{attribute 'linkalways'} 
{attribute 'no_explicit_call' := 'This FB is a CLASS and must be accessed using methods or properties'}
{attribute 'enable_dynamic_creation'}
FUNCTION_BLOCK _ETcVnWorldCoordinateSystem EXTENDS EnumDatatypeBase
VAR
	localData : ETcVnWorldCoordinateSystem;
	activeData : REFERENCE TO ETcVnWorldCoordinateSystem;
	enumBaseDatatype : _DINT(localData);
END_VAR

METHOD PRIVATE AddLocalEnumeration
VAR_INPUT
	Enumeration : T_MAXSTRING;
	Value : ETcVnWorldCoordinateSystem;
END_VAR
AddEnumeration(Enumeration, Value);
END_METHOD

PROPERTY PUBLIC Address : PVOID
GET
Address := ADR(activeData);
END_GET
END_PROPERTY

METHOD PUBLIC ClearReference
VAR_INPUT
END_VAR
activeData REF= localData;
SetBaseDatatypeReference();
END_METHOD

METHOD PUBLIC Clone : I_Datatype
VAR
    pClone : POINTER TO _ETcVnWorldCoordinateSystem;
END_VAR
pClone := __NEW(_ETcVnWorldCoordinateSystem(InitialValue := Value));
Clone := pClone^;
END_METHOD

METHOD FB_init : BOOL
VAR_INPUT
	bInitRetains : BOOL; // if TRUE, the retain variables are initialized (warm start / cold start)
	bInCopyCode : BOOL;  // if TRUE, the instance afterwards gets moved into the copy code (online change)
	InitialValue : ETcVnWorldCoordinateSystem;
END_VAR
localData := InitialValue;
AddBaseDatatype(enumBaseDatatype);
ClearReference();

AddLocalEnumeration('TCVN_WCS_X_RIGHT_Y_DOWN' , ETcVnWorldCoordinateSystem.TCVN_WCS_X_RIGHT_Y_DOWN);
AddLocalEnumeration('TCVN_WCS_X_DOWN_Y_RIGHT', ETcVnWorldCoordinateSystem.TCVN_WCS_X_DOWN_Y_RIGHT);
AddLocalEnumeration('TCVN_WCS_X_LEFT_Y_DOWN', ETcVnWorldCoordinateSystem.TCVN_WCS_X_LEFT_Y_DOWN);
AddLocalEnumeration('TCVN_WCS_X_UP_Y_RIGHT', ETcVnWorldCoordinateSystem.TCVN_WCS_X_UP_Y_RIGHT);
AddLocalEnumeration('TCVN_WCS_X_RIGHT_Y_UP', ETcVnWorldCoordinateSystem.TCVN_WCS_X_RIGHT_Y_UP);
AddLocalEnumeration('TCVN_WCS_X_DOWN_Y_LEFT', ETcVnWorldCoordinateSystem.TCVN_WCS_X_DOWN_Y_LEFT);
AddLocalEnumeration('TCVN_WCS_X_LEFT_Y_UP', ETcVnWorldCoordinateSystem.TCVN_WCS_X_LEFT_Y_UP);
AddLocalEnumeration('TCVN_WCS_X_UP_Y_LEFT', ETcVnWorldCoordinateSystem.TCVN_WCS_X_UP_Y_LEFT);
END_METHOD

PROPERTY PUBLIC Identifier : T_MAXSTRING
GET
Identifier := 'ETcVnWorldCoordinateSystem';
END_GET
END_PROPERTY

METHOD IsEnumeratorValueEqual : BOOL
VAR_INPUT
	Enumerator : I_KeyValueForwardEnumerator;
END_VAR
VAR
	storedValue : ETcVnWorldCoordinateSystem;
END_VAR
IF NOT Enumerator.TryGet(storedValue) THEN
	RETURN;
END_IF

IsEnumeratorValueEqual := storedValue = activeData;
END_METHOD

METHOD PUBLIC MakeReferenceTo
VAR_INPUT
	ReferenceTarget : REFERENCE TO ETcVnWorldCoordinateSystem;
END_VAR
activeData REF= ReferenceTarget;
SetBaseDatatypeReference();
END_METHOD

METHOD PROTECTED SetBaseDatatypeReference
VAR_INPUT
END_VAR
enumBaseDatatype.MakeReferenceTo(activeData);
END_METHOD

PROPERTY PUBLIC Size : UDINT
GET
Size := SIZEOF(activeData);
END_GET
END_PROPERTY

METHOD TryMakeReferenceTo : BOOL
VAR_INPUT
	Target : I_Datatype;
END_VAR
VAR
	pTargetData : POINTER TO ETcVnWorldCoordinateSystem;
END_VAR
IF NOT IsEquivalentTo(Target) THEN
	RETURN;
END_IF

pTargetData := Target.Address;
activeData REF= pTargetData^;
SetBaseDatatypeReference();
TryMakeReferenceTo := TRUE;
END_METHOD

PROPERTY PUBLIC Value : ETcVnWorldCoordinateSystem
GET
Value := activeData;
END_GET
SET
activeData := Value;
END_SET
END_PROPERTY

END_FUNCTION_BLOCK

(* stored: Version 1.1.0.1, ProductVersion 3.1.4024.13
   POU _ETcVnWorldCoordinateSystem: Id {235e61e2-5d3d-043c-262e-e83edc5adb14}, SpecialFunc None
   Folder Core: Id {d6405b57-d99a-02a6-31c7-c060a403458b}
   Folder Protected: Id {fe40e79b-4cec-0bcd-0cc8-45e727329045}
   Folder Customize: Id {33fe7baf-cb5d-0759-23df-f0978ef822f8}
   Folder Constructor: Id {bb911ded-345e-03e7-2696-8eaf38f3a321}
   Folder Private: Id {a1382847-d034-03ca-3fc7-e535256b42dd}
   Folder Protected: Id {205802c8-b1d5-0cc0-0a49-c2a9fb111632}
   Method AddLocalEnumeration: Id {5c86a2d5-30c6-0385-36b6-ecbe6a3bf5eb}
   Property Address: Id {c859675d-928d-0eb8-0079-4ff989b745be}
   Get Get: Id {b533b12b-97f4-0ca6-0f99-e117360cad6f}
   Method ClearReference: Id {976e8571-8f50-0787-26af-3912f8797dd4}
   Method Clone: Id {767cf40d-300b-0e3d-2f8b-3d0a349f4f77}
   Method FB_init: Id {02033452-19a0-0ea9-1749-296e9cdf01be}
   Property Identifier: Id {d50350db-e945-08ff-1686-0b3d17a3a989}
   Get Get: Id {9c0128e5-06a4-01db-0b79-e492c435f246}
   Method IsEnumeratorValueEqual: Id {8e91c633-cea1-075b-3387-8823156b512c}
   Method MakeReferenceTo: Id {14579730-ceda-00a4-135e-8db8796c2903}
   Method SetBaseDatatypeReference: Id {40fe89d9-ca4d-0800-276d-aef03ed957c3}
   Property Size: Id {cb9fa0c1-3773-0286-0016-534eda4e8ea4}
   Get Get: Id {35c30f9a-d7c4-03ed-045a-4d05804389b9}
   Method TryMakeReferenceTo: Id {c755a6eb-b986-0538-1127-77d825663004}
   Property Value: Id {61605790-b832-02a7-1c20-95353ba766d2}
   Get Get: Id {1c6427ea-037e-030b-3ce4-17be0c45350f}
   Set Set: Id {53a134b2-20e4-0afe-014f-709ae28b2314} *)
